Omron CX-Programmer project  (CX-Programmer ?)

# PLC :  

## Function block Humidity
VAR_INPUT
  Current_Value_Humidity : INT;
END_VAR
VAR_OUTPUT
  Humidity : REAL;
END_VAR
VAR
  IHumid : REAL;
  Real_Value_Humidity : REAL;
END_VAR
Real_Value_Humidity:= INT_TO_REAL(Current_Value_Humidity);
IHumid:= (Real_Value_Humidity/250.0)+4.0;
Humidity:= (IHumid-4.0)/16.0*95.0;

## Function block Temperature
VAR_INPUT
  Current_Value : INT;
END_VAR
VAR_OUTPUT
  Temp : REAL;
END_VAR
VAR
  Itemp : REAL;
  Real_Current_Value : REAL;
END_VAR
Real_Current_Value:= INT_TO_REAL(Current_Value);
Itemp:= 4.0 + (Real_Current_Value / 4000.0) * 16.0;
Temp:= ((Itemp-4.0)/16.0)*90.0-20.0;